(* IEC 61131-3 sources: llm-plc-st-eval/data/processed_definitivo/qwen2.5-coder_14b/C6/zero_shot, 1 file *)

(* ---- ejec_1.st ---- *)
VAR
        enfriadorEstado : BOOL := FALSE;
    END_VAR

    IF tempC >= 80.0 THEN
        enfriador := TRUE;
        enfriadorEstado := TRUE;
    ELSIF tempC < 75.0 THEN
        enfriador := FALSE;
        enfriadorEstado := FALSE;
    ELSE
        enfriador := enfriadorEstado;
    END_IF
